(* IEC 61131-3 sources: llm-plc-st-eval/data/definitivo/gpt-4o-2024-08-06/B1/few_shot, 3 files *)

(* ---- ejec_1.st ---- *)
```pascal
FUNCTION_BLOCK FB_Motor
VAR_INPUT
    btnMarcha : BOOL; (* Botón de marcha *)
    btnParo : BOOL;   (* Botón de paro *)
    btnEmerg : BOOL;  (* Botón de paro de emergencia *)
END_VAR
VAR_OUTPUT
    motorOn : BOOL;   (* Estado del motor *)
END_VAR
VAR
    estadoMotor : BOOL; (* Estado interno del motor *)
END_VAR

(* Lógica de control del motor *)
IF btnEmerg THEN
    estadoMotor := FALSE; (* Paro de emergencia, motor apagado *)
ELSIF btnParo THEN
    estadoMotor := FALSE; (* Botón de paro, motor apagado *)
ELSIF btnMarcha THEN
    estadoMotor := TRUE;  (* Botón de marcha, motor encendido *)
END_IF

motorOn := estadoMotor; (* Salida del estado del motor *)
END_FUNCTION_BLOCK
```

(* ---- ejec_2.st ---- *)
```pascal
FUNCTION_BLOCK FB_Motor
VAR_INPUT
    btnMarcha : BOOL; (* Boton de marcha *)
    btnParo : BOOL;   (* Boton de paro *)
    btnEmerg : BOOL;  (* Boton de paro de emergencia *)
END_VAR
VAR_OUTPUT
    motorOn : BOOL;   (* Estado del motor *)
END_VAR
VAR
    motorLatch : BOOL; (* Latch para mantener el motor encendido *)
END_VAR

(* Control de arranque y paro del motor *)
IF btnEmerg THEN
    (* Si se activa el paro de emergencia, el motor se apaga y no puede rearrancar *)
    motorLatch := FALSE;
ELSIF btnParo THEN
    (* Si se pulsa el boton de paro, el motor se apaga *)
    motorLatch := FALSE;
ELSIF btnMarcha THEN
    (* Si se pulsa el boton de marcha, el motor se enciende y se mantiene encendido *)
    motorLatch := TRUE;
END_IF

(* Actualizar el estado del motor *)
motorOn := motorLatch;
END_FUNCTION_BLOCK
```

(* ---- ejec_3.st ---- *)
```pascal
FUNCTION_BLOCK FB_Motor
VAR_INPUT
    btnMarcha : BOOL; (* Botón de marcha *)
    btnParo : BOOL;   (* Botón de paro *)
    btnEmerg : BOOL;  (* Botón de paro de emergencia *)
END_VAR
VAR_OUTPUT
    motorOn : BOOL;   (* Estado del motor *)
END_VAR
VAR
    estadoMotor : BOOL; (* Estado interno del motor *)
END_VAR

(* Control de arranque y paro del motor *)
IF btnEmerg THEN
    estadoMotor := FALSE; (* Paro de emergencia, motor apagado *)
ELSIF btnParo THEN
    estadoMotor := FALSE; (* Botón de paro, motor apagado *)
ELSIF btnMarcha THEN
    estadoMotor := TRUE;  (* Botón de marcha, motor encendido *)
END_IF

motorOn := estadoMotor; (* Salida del estado del motor *)
END_FUNCTION_BLOCK
```
